KUKA KRL program: JointTargets.src

&ACCESS RVP
&REL 1
&PARAM TEMPLATE = C:\KRC\Roboter\Template\vorgabe
&PARAM EDITMASK = *
DEF JointTargets ( )


; GLOBAL INTERRUPT DECL 3 WHEN $STOPMESS==TRUE DO IR_STOPM ( )
; INTERRUPT ON 3

;FOLD Initialise and set default speed
BAS (#INITMOV,0)
BAS (#VEL_PTP,100)
BAS (#ACC_PTP,20)
$VEL.CP=0.2
BAS (#TOOL,0)
BAS (#BASE,0)
;ENDFOLD

;;FOLD STARTPOS
;$BWDSTART = FALSE
;PDAT_ACT = PDEFAULT
;BAS(#PTP_DAT)
;FDAT_ACT = {TOOL_NO 0,BASE_NO 0,IPO_FRAME #BASE}
;BAS(#FRAMES)
;;ENDFOLD

$ADVANCE = 5

;FOLD ---- Quickly skip BCO ----
; PTP $AXIS_ACT
;ENDFOLD

;FOLD ---- GO HOME ----
; PTP {A1 0.000, A2 -90.000, A3 90.000, A4 0.000, A5 0.000, A6 0.000, E1 0, E2 0, E3 0, E4 0, E5 0, E6 0}
;ENDFOLD


; Program generated by VerticalBot Studio for KUKA KR 6 R900 sixx on 25/10/2026 12:00:00
; Using nominal kinematics.
; ---- Setting reference (Base) ----
; BASE_DATA[2] = {FRAME: X 100.000,Y -50.000,Z 20.000,A 30.000,B 0.000,C 0.000}
$BASE = {FRAME: X 100.000,Y -50.000,Z 20.000,A 30.000,B 0.000,C 0.000}
; $BASE = BASE_DATA[2]
; --------------------------
; ---- Setting tool (TCP) ----
; TOOL_DATA[1] = {FRAME: X 10.000,Y 0.000,Z 120.000,A 0.000,B 15.000,C 0.000}
$TOOL = {FRAME: X 10.000,Y 0.000,Z 120.000,A 0.000,B 15.000,C 0.000}
; $TOOL = TOOL_DATA[1]
; --------------------------
PTP {A1 10.00000,A2 -80.00000,A3 100.00000,A4 20.00000,A5 40.00000,A6 -30.00000}
; Linear movement using joint targets is not supported. Change the target type to cartesian or use a joint movement.
PTP {A1 18.00000,A2 -76.00000,A3 100.00000,A4 20.00000,A5 40.00000,A6 -30.00000}
LIN {X 521.453,Y -74.708,Z 545.847,A 177.940,B 18.811,C 176.970}
; Linear movement using joint targets is not supported. Change the target type to cartesian or use a joint movement.
$APO.CPTP = 5
$APO.CDIS = 5.000
PTP {A1 10.00000,A2 -80.00000,A3 100.00000,A4 20.00000,A5 40.00000,A6 -30.00000} C_PTP
; Linear movement using joint targets is not supported. Change the target type to cartesian or use a joint movement.
PTP {A1 18.00000,A2 -76.00000,A3 100.00000,A4 20.00000,A5 40.00000,A6 -30.00000} C_PTP
LIN {X 521.453,Y -74.708,Z 545.847,A 177.940,B 18.811,C 176.970} C_DIS
; Linear movement using joint targets is not supported. Change the target type to cartesian or use a joint movement.
PTP {A1 10.00000,A2 -80.00000,A3 100.00000,A4 20.00000,A5 40.00000,A6 -30.00000}
END
